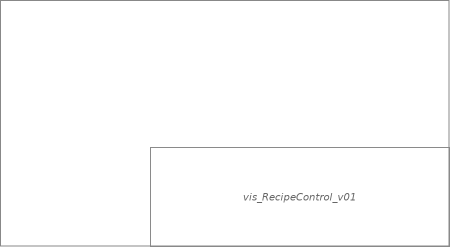
VISUALIZATION vis_RecipeTest  // 450x247
    Frame (150,147 300x100)
        shows vis_RecipeControl_v01(Definition := 'R_Open1')
END_VISUALIZATION

(* stored: Version 1.1.0.1, ProductVersion 3.1.4024.12
   Visu vis_RecipeTest: Id {ed879417-48d7-430b-ba4a-27e7b64a7d12} *)
